// TIA Portal V21 export
VAR_GLOBAL   // PLC tag table "Reset"
   reset AT %I5.7 : Bool;
   reset_led AT %Q1.7 : Bool;
END_VAR
